Staubli VAL3: setBtnColor.pgx

public program setBtnColor(num x_nJogmode)
  local string l_sNULLcolor
  local num l_i
  local string l_sbtn
  local string l_sSELcolor
begin
  l_sNULLcolor="#FFFFFF"
  l_sSELcolor="#3399FF"

  switch x_nJogmode
    case 0
      for l_i = 1 to 4 step 1
        l_sbtn="btn"+toString("",l_i)
        userPageSet("jogmode",l_sbtn,"style.backgroundColor",l_sNULLcolor)
      endFor
    break
    case 1
      userPageSet("jogmode","btn1","style.backgroundColor",l_sNULLcolor)
      userPageSet("jogmode","btn2","style.backgroundColor",l_sSELcolor)
      userPageSet("jogmode","btn3","style.backgroundColor",l_sNULLcolor)
      userPageSet("jogmode","btn4","style.backgroundColor",l_sNULLcolor)
    break
    case 2
      userPageSet("jogmode","btn1","style.backgroundColor",l_sNULLcolor)
      userPageSet("jogmode","btn3","style.backgroundColor",l_sSELcolor)
      userPageSet("jogmode","btn2","style.backgroundColor",l_sNULLcolor)
      userPageSet("jogmode","btn4","style.backgroundColor",l_sNULLcolor)
    break
    case 3
      userPageSet("jogmode","btn1","style.backgroundColor",l_sNULLcolor)
      userPageSet("jogmode","btn2","style.backgroundColor",l_sNULLcolor)
      userPageSet("jogmode","btn3","style.backgroundColor",l_sNULLcolor)
      userPageSet("jogmode","btn4","style.backgroundColor",l_sSELcolor)
    break

  endSwitch
end
